(* PLC project Unnamed, Unknown Unnamed 1 *)
(* stored: creationDateTime 2023-10-17T07:56:28, modificationDateTime 2023-10-17T10:02:17 *)

PROGRAM plc1
  VAR
    ColorSensor_RED AT %IW0 : INT;
    ColorSensor_GREEN AT %IW1 : INT;
    ColorSensor_BLUE AT %IW2 : INT;
    RangeSensor AT %IW3 : INT;
    Pump AT %QX0.4 : BOOL := False;
    treatmentComplete AT %IX100.0 : BOOL := False;  (* Value received from PLC2 *)
  END_VAR
  VAR
    desiredDistanceFill : REAL := 7.0;
    measuredDistance : REAL;
  END_VAR

            
(*Workaround to distance measure bug*)
measuredDistance := INT_TO_REAL(RangeSensor)/100.0;
desiredDistanceFill := 7.0;

IF treatmentComplete THEN
        IF measuredDistance > desiredDistanceFill THEN
          Pump := TRUE;
        ELSE
          Pump := FALSE;
        END_IF;
END_IF;
          
END_PROGRAM

CONFIGURATION Config0
  RESOURCE Res0 ON PLC
    TASK task0(INTERVAL := T#20ms, PRIORITY := 0);
    PROGRAM instance0 WITH task0 : plc1;
  END_RESOURCE
END_CONFIGURATION
